// TIA Portal V20 export
// export: Created 2026-10-11T05:25:31.2300143Z, ExportSetting WithDefaults, DisplayName Totally Integrated Automation Portal, DisplayVersion V20, DisplayName TIA Portal Openness, DisplayVersion V20, DisplayName TIA Portal Teamcenter Gateway, DisplayVersion V20, DisplayName TIA Portal Version Control Interface, DisplayVersion V20, DisplayName SINAMICS Startdrive Advanced, DisplayVersion V20 SP1 Update 2, DisplayName SINAMICS Startdrive G110M, G120, G120C, G120D, G120P, G115D, DisplayVersion V20 SP1 Update 2, DisplayName SINAMICS Startdrive G130, G150, S120, S150, SINAMICS MV, G220, S200, S210, DisplayVersion V20 SP1 Update 2, DisplayName STEP 7 Professional, DisplayVersion V20, DisplayName STEP 7 Safety, DisplayVersion V20, DisplayName WinCC Basic/Comfort/Advanced, DisplayVersion V20, DisplayName WinCC Professional, DisplayVersion V20, DisplayName WinCC Unified, DisplayVersion V20
FUNCTION "FRK_ManualApply" : Void   // FC57, SCL
{ S7_Optimized_Access := 'TRUE' }
VERSION : 0.1
// stored: AutoNumber true, IsIECCheckEnabled false, SetENOAutomatically false, UDAEnableTagReadback false
   VAR_INPUT
      Request : "ST_HmiRequest";
      Status : "ST_ModuleStatus";
      Core : "FRK_Core";
      Commands : Array[1..12] of "ST_CommandInfo";
      Count : DInt;
      Conditions : Array[1..16] of "FRK_ManualConditionRow";
   END_VAR
   VAR_IN_OUT
      Report : "ST_ReleaseReport";
      Execute : Bool;
      Command : DInt;
      ManualOwned : Bool;
   END_VAR
   VAR_TEMP
      Index : Int;
      Supported : Bool;
      PreviousCount : Int;
   END_VAR
BEGIN

   #Supported := FALSE;
   IF #Count >= 0 AND #Count <= 12 THEN
       FOR #Index := 1 TO DINT_TO_INT(#Count) DO
           IF #Commands[#Index].Value = #Request.IntValue AND #Commands[#Index].Style = 0 THEN
               #Supported := TRUE;
           END_IF;
       END_FOR;
   END_IF;
   IF NOT #Supported THEN
       "FRK_ReleaseReason"(Report := #Report,
                           Description := WSTRING#'std.error.unsupportedHmiRequest',
                           Reason := 2008,
                           Path := STRING_TO_WSTRING(#Status.Name),
                           Kind := 4);
   END_IF;
   IF #Core.Exec <> 0 OR #Execute OR #Core.ReleasePending THEN
       "FRK_ReleaseReason"(Report := #Report,
                           Description := WSTRING#'std.error.hmiRequestRejected',
                           Reason := 2011,
                           Path := STRING_TO_WSTRING(#Status.Name),
                           Kind := 4);
   END_IF;
   FOR #Index := 1 TO 16 DO
       IF #Conditions[#Index].Used AND NOT #Conditions[#Index].Ok THEN
           IF #Conditions[#Index].Value = 0 OR #Conditions[#Index].Value = #Request.IntValue THEN
               #PreviousCount := #Report.Count;
               "FRK_ReleaseReason"(Report := #Report,
                                   Description := #Conditions[#Index].Diag.Description,
                                   Reason := #Conditions[#Index].Diag.ReasonCode,
                                   Path := STRING_TO_WSTRING(#Status.Name),
                                   Kind := 3);
               IF #Report.Count > #PreviousCount THEN
                   #Report.Reasons[#Report.Count].Bypassable := #Conditions[#Index].Bypassable;
               END_IF;
           END_IF;
       END_IF;
   END_FOR;
   IF #Request.Kind = 11 AND #Report.Released THEN
       #Command := #Request.IntValue;
       #Execute := TRUE;
       #ManualOwned := TRUE;
   END_IF;
END_FUNCTION
